Fanuc KAREL source: kt00533.KL

-- PROVISIONAL review KL for V770-1; original PC SHA256 14fe9609ac2c8dda611e6b5799024987a39600cf6079b06dce537048a9321325
-- Incomplete behavior may be omitted. Consult companion uncertainty JSON. Do not deploy.
PROGRAM KT00533
%NOLOCKGROUP
VAR
  OUT : BOOLEAN
-- UNRESOLVED_DECL P1 type=000199
-- UNRESOLVED_DECL P2 type=000101
BEGIN
  -- UNRESOLVED_PC offsets 5-33; opcodes 49,7E,49,AC,23
  -- UNRESOLVED_PC offsets 38-42; opcodes 7F
END KT00533
